(* IEC 61131-3 sources: LASAL/Network/EncoderSimulation, 1 file *)

(* ---- ONE_EncoderSimulation_Table.st ---- *)
#define OBJECTS_CONFIG

FUNCTION GLOBAL TAB ONE_EncoderSimulation
-1$UINT, 0$UINT,
0$UINT, 0$UINT,

1$UDINT,
TO_UDINT(1540101447), "Encoders", 0$UINT, 0$UINT, 1$UINT,

_NO_ATTR, TO_UDINT(1799354257), "ENCODERS1",

//Internal connections
0$UDINT,
0$UDINT,
0$UDINT,
0$UDINT,

//Initialization values
0$UDINT,
8$UDINT,
TO_UDINT(0), "KV", TO_UDINT(100),//|EncoderSimulation.Encoders1.KV;
TO_UDINT(0), "MUL", TO_UDINT(11700),//|EncoderSimulation.Encoders1.MUL;
TO_UDINT(0), "DIV", TO_UDINT(1000),//|EncoderSimulation.Encoders1.DIV;
TO_UDINT(0), "InvertOutput", TO_UDINT(1),//|EncoderSimulation.Encoders1.InvertOutput;
TO_UDINT(0), "pos_in_fixed", TO_UDINT(-1),//|EncoderSimulation.Encoders1.pos_in_fixed;
TO_UDINT(0), "pos_in_steppermotor", TO_UDINT(0),//|EncoderSimulation.Encoders1.pos_in_steppermotor;
TO_UDINT(0), "Speed_out", TO_UDINT(0),//|EncoderSimulation.Encoders1.Speed_out;
TO_UDINT(0), "Pos_out", TO_UDINT(-1),//|EncoderSimulation.Encoders1.Pos_out;

//Symbolic initialization values
0$UDINT,
0$UDINT,

//Initialization of string values
0$UDINT,
0$UDINT,

//Configuration of tasks (RealTime, Cyclic, Background)
0$UDINT,
1$UDINT,
TO_UDINT(0), (1)$UDINT, 4194306$DINT, 	//ENCODERS1

0$UDINT,
0$UDINT,

0$UDINT,
0$UDINT,

//External connections
0$UDINT,
4$UDINT,
TO_UDINT(0), "pos_in_fixed", C_DIR, TO_UDINT(3024798335), "ST0111","Encoder",
TO_UDINT(0), "pos_in_steppermotor", C_DIR, TO_UDINT(201264582), "ST1511","ActPosition",
TO_UDINT(0), "Speed_out", C_DIR, TO_UDINT(3024798335), "ST0111","FreqOut",
TO_UDINT(0), "Pos_out", C_DIR, TO_UDINT(3024798335), "ST0111","ClockCounter",

//Magic internal connections
0$UDINT,
0$UDINT,

//Configuration of timeslots of tasks (RealTime, Cyclic)
#ifdef __LSLLDR_TIMESLOTS__
0$UDINT,
0$UDINT,

0$UDINT,
0$UDINT,

#endif //__LSLLDR_TIMESLOTS__

//MultiMaster connections
#ifdef __LSLLDR_MULTIMASTER__
0$UDINT,
0$UDINT,
#endif //__LSLLDR_MULTIMASTER__

//Configuration for task ID (RealTime, CyclicTime)
#ifdef __LSLLDR_TASKID__
"\\\\TASKS2  "
0$UDINT,
1$UDINT,
(0)$UDINT, 	//ENCODERS1

0$UDINT,
0$UDINT,

0$UDINT,
0$UDINT,

#endif //__LSLLDR_TASKID__

END_FUNCTION
